FUNCTION_BLOCK CustomStopActuator (* Basic Function Block Type *)
  (* Standard: 61499-2 *)
  (* Version 0.0, 7/2/2026, Template *)
  PACKAGE Main;
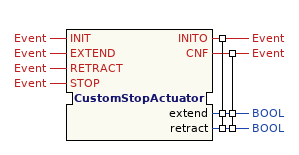
  EVENT_INPUT
    INIT; (* Initialization Request *)
    EXTEND; (* Normal Execution Request *)
    RETRACT;
    STOP;
  END_EVENT
  EVENT_OUTPUT
    INITO WITH extend, retract; (* Initialization Confirm *)
    CNF WITH extend, retract; (* Execution Confirmation *)
  END_EVENT
  VAR_OUTPUT
    extend : BOOL; (* Output event qualifier *)
    retract : BOOL;
  END_VAR
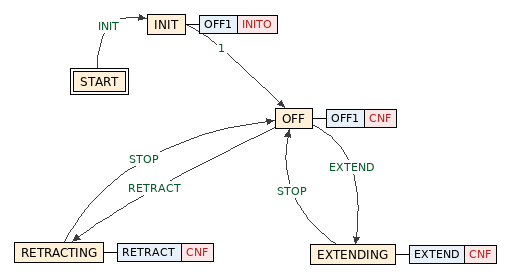
  EC_STATES
    START; (* Initial State *)
    INIT : OFF1 -> INITO; (* Initialization *)
    OFF : OFF1 -> CNF;
    EXTENDING : EXTEND -> CNF;
    RETRACTING : RETRACT -> CNF;
  END_STATES
  EC_TRANSITIONS
    START TO INIT := INIT;
    INIT TO OFF := 1;
    OFF TO RETRACTING := RETRACT;
    RETRACTING TO OFF := STOP;
    OFF TO EXTENDING := EXTEND;
    EXTENDING TO OFF := STOP;
  END_TRANSITIONS
  ALGORITHM INIT IN ST: (* Initialization algorithm *)
;
  END_ALGORITHM
  ALGORITHM REQ IN ST: (* Normally executed algorithm *)
;
  END_ALGORITHM
  ALGORITHM OFF1 IN ST:
extend := FALSE;
retract := FALSE;
  END_ALGORITHM
  ALGORITHM EXTEND IN ST:
extend := TRUE;
retract := FALSE;
  END_ALGORITHM
  ALGORITHM RETRACT IN ST:
extend := FALSE;
retract := TRUE;
  END_ALGORITHM
END_FUNCTION_BLOCK
